(* IEC 61131-3 sources: RootPLC/conformance/cases/lexical, 40 files *)

(* ---- warn_soft_keyword_name.st ---- *)
(* spec: [lexical.keywords.soft]
   expect: warning RP0124
   run: PRG_Main cycles=2
   assert: n = 2
   assert: lit = TRUE *)
FUNCTION_BLOCK FB_Sequence
VAR_INPUT
    Step : INT;
    On : BOOL;
END_VAR
VAR_OUTPUT
    Task : DINT;
END_VAR
CASE Step OF
    1: Task := Task + 1;
END_CASE;
END_FUNCTION_BLOCK

PROGRAM PRG_Main
VAR
    seq : FB_Sequence;
    n : DINT;
    lit : BOOL;
    lamp AT %QX0.0 : BOOL;
END_VAR
seq(Step := 1, On := TRUE);
n := seq.Task;
lamp := seq.On;
lit := lamp;
END_PROGRAM

(* ---- err_bad_based_digit.st ---- *)
(* spec: [lexical.literal.integer]
   expect: error RP0008 *)
PROGRAM PRG_Main
VAR
    x : INT := 8#19;
END_VAR

END_PROGRAM

(* ---- err_bad_escape.st ---- *)
(* spec: [lexical.literal.escape]
   expect: error RP0010 *)
PROGRAM PRG_Main
VAR
    s : STRING := 'a$Qb';
END_VAR

END_PROGRAM

(* ---- err_char_two.st ---- *)
(* spec: [lexical.literal.char]
   expect: error RP0008 *)
PROGRAM PRG_Main
VAR
    c : CHAR := CHAR#'ab';
END_VAR

END_PROGRAM

(* ---- err_date_invalid.st ---- *)
(* spec: [lexical.literal.date]
   expect: error RP0012 *)
PROGRAM PRG_Main
VAR
    d : DATE := D#2026-02-30;
END_VAR

END_PROGRAM

(* ---- err_direct_variable.st ---- *)
(* spec: [lexical.direct-variable]
   expect: error RP0016 *)
PROGRAM PRG_Main
VAR
    x AT %IZ0 : BOOL;
END_VAR

END_PROGRAM

(* ---- err_duration_fraction_not_last.st ---- *)
(* spec: [lexical.literal.duration]
   expect: error RP0011 *)
PROGRAM PRG_Main
VAR
    t : TIME := T#1.5s20ms;
END_VAR

END_PROGRAM

(* ---- err_duration_order.st ---- *)
(* spec: [lexical.literal.duration]
   expect: error RP0011 *)
PROGRAM PRG_Main
VAR
    t : TIME := T#5s1m;
END_VAR

END_PROGRAM

(* ---- err_invalid_char.st ---- *)
(* spec: [lexical.source.charset] [lexical.punctuation]
   expect: error RP0005 *)
PROGRAM PRG_Main
VAR
    x : INT;
END_VAR
x := 1 @ 2;
END_PROGRAM

(* ---- err_keyword_identifier.st ---- *)
(* spec: [lexical.keyword]
   expect: error RP0004 *)
PROGRAM PRG_Main
VAR
    end_if : INT;
END_VAR

END_PROGRAM

(* ---- err_non_ascii_identifier.st ---- *)
(* spec: [lexical.source.charset]
   expect: error RP0005 *)
PROGRAM PRG_Main
VAR
    温度 : INT;
END_VAR

END_PROGRAM

(* ---- err_real_no_fraction.st ---- *)
(* spec: [lexical.literal.real]
   expect: error RP0008 *)
PROGRAM PRG_Main
VAR
    x : LREAL := 1.;
END_VAR

END_PROGRAM

(* ---- err_string_latin1.st ---- *)
(* spec: [lexical.literal.string.latin1]
   expect: error RP0009 *)
PROGRAM PRG_Main
VAR
    s : STRING := '温度';
END_VAR

END_PROGRAM

(* ---- err_tod_hour24.st ---- *)
(* spec: [lexical.literal.date]
   expect: error RP0012 *)
PROGRAM PRG_Main
VAR
    t : TOD := TOD#24:00:00;
END_VAR

END_PROGRAM

(* ---- err_typed_unknown.st ---- *)
(* spec: [lexical.literal.typed]
   expect: error RP0014 *)
PROGRAM PRG_Main
VAR
    x : INT := FOO#5;
END_VAR

END_PROGRAM

(* ---- err_underscore_double.st ---- *)
(* spec: [lexical.literal.underscore]
   expect: error RP0007 *)
PROGRAM PRG_Main
VAR
    x : INT := 1__0;
END_VAR

END_PROGRAM

(* ---- err_underscore_trailing.st ---- *)
(* spec: [lexical.literal.underscore]
   expect: error RP0007 *)
PROGRAM PRG_Main
VAR
    x : INT := 100_;
END_VAR

END_PROGRAM

(* ---- err_unterminated_comment.st ---- *)
(* spec: [lexical.comment.unterminated]
   expect: error RP0001 *)
PROGRAM PRG_Main (* never closed
END_PROGRAM

(* ---- err_unterminated_pragma.st ---- *)
(* spec: [lexical.pragma]
   expect: error RP0015 *)
PROGRAM PRG_Main
{attribute 'hide'
END_PROGRAM

(* ---- err_unterminated_string.st ---- *)
(* spec: [lexical.literal.string]
   expect: error RP0002 *)
PROGRAM PRG_Main
VAR
    s : STRING := 'abc
    n : INT;
END_VAR

END_PROGRAM

(* ---- ok_char_literals.st ---- *)
(* spec: [lexical.literal.char]
   expect: ok
   run: PRG_Main cycles=1
   assert: c = CHAR#'a' *)
PROGRAM PRG_Main
VAR
    c : CHAR := CHAR#'a';
    w : WCHAR := WCHAR#"b";
END_VAR

END_PROGRAM

(* ---- ok_comments.st ---- *)
(* spec: [lexical.comment.block] [lexical.comment.cblock] [lexical.comment.line] [lexical.whitespace] [lexical.source.encoding]
   expect: ok
   run: PRG_Main cycles=1
   assert: s = '/* not a comment */'
   assert: n = 1 *)
PROGRAM PRG_Main
VAR
    s : STRING := '/* not a comment */'; // line comment
    s2 : STRING := '(* not a comment *)';
	n : INT; /* C-style */
END_VAR
(* block
   comment *)
n := 1;
END_PROGRAM

(* ---- ok_date_literals.st ---- *)
(* spec: [lexical.literal.date]
   expect: ok *)
PROGRAM PRG_Main
VAR
    d : DATE := D#2026-11-03;
    t_day : TOD := TOD#14:30:00.5;
    stamp : DT := DT#2026-11-03-14:30:00;
    ld : LDATE := LDATE#2024-02-29;
END_VAR

END_PROGRAM

(* ---- ok_direct_variable.st ---- *)
(* spec: [lexical.direct-variable]
   expect: ok *)
PROGRAM PRG_Main
VAR
    start_btn AT %IX0.0 : BOOL;
    lamp AT %QX0.1 : BOOL;
    level AT %IW2 : WORD;
    spare AT %I* : BOOL;
END_VAR

END_PROGRAM

(* ---- ok_duration_literals.st ---- *)
(* spec: [lexical.literal.duration]
   expect: ok
   run: PRG_Main cycles=1
   assert: t1 = T#90m
   assert: t3 = T#1500ms *)
PROGRAM PRG_Main
VAR
    t1 : TIME := T#1h_30m;
    t2 : TIME := T#90m;
    t3 : TIME := T#1.5s;
    t4 : LTIME := LTIME#5us;
    t5 : TIME := t#-250ms;
END_VAR

END_PROGRAM

(* ---- ok_identifier_case.st ---- *)
(* spec: [lexical.identifier] [lexical.identifier.case]
   expect: ok
   run: PRG_Main cycles=1
   assert: motor_on = TRUE
   assert: _x1 = 3 *)
PROGRAM PRG_Main
VAR
    Motor_On : BOOL;
    _x1 : INT;
END_VAR
MOTOR_ON := TRUE;
_X1 := 3;
END_PROGRAM

(* ---- ok_integer_literals.st ---- *)
(* spec: [lexical.literal.integer] [lexical.literal.underscore] [lexical.literal.sign]
   expect: ok
   run: PRG_Main cycles=1
   assert: a = 1000000
   assert: b = 165
   assert: c = 15
   assert: d = 255
   assert: e = -128 *)
PROGRAM PRG_Main
VAR
    a : DINT := 1_000_000;
    b : INT := 2#1010_0101;
    c : INT := 8#17;
    d : DINT := 16#ff;
    e : SINT := -128;
END_VAR

END_PROGRAM

(* ---- ok_longest_match.st ---- *)
(* spec: [lexical.longest-match] [lexical.punctuation] [types.derived.array]
   expect: ok
   run: PRG_Main cycles=1
   assert: b = TRUE
   assert: a[10] = 1 *)
PROGRAM PRG_Main
VAR
    a : ARRAY[1..10] OF INT;
    x : INT := 1;
    y : INT := 2;
    b : BOOL;
END_VAR
b := x<=y;
a[10] := x**2;
END_PROGRAM

(* ---- ok_pragma_attribute.st ---- *)
(* spec: [lexical.pragma]
   expect: ok *)
PROGRAM PRG_Main
VAR
    {attribute 'hide'}
    x : INT;
END_VAR

END_PROGRAM

(* ---- ok_real_literals.st ---- *)
(* spec: [lexical.literal.real]
   expect: ok
   run: PRG_Main cycles=1
   assert: r = 1500.0
   assert: s = 0.25
   assert: t = 0.01 *)
PROGRAM PRG_Main
VAR
    r : LREAL := 1.5E3;
    s : REAL := 0.25;
    t : LREAL := 1.0e-2;
END_VAR

END_PROGRAM

(* ---- ok_strings.st ---- *)
(* spec: [lexical.literal.string] [lexical.literal.escape]
   expect: ok
   run: PRG_Main cycles=1
   assert: h = 'A' *)
PROGRAM PRG_Main
VAR
    s : STRING := 'it$'s $$5$N';
    w : WSTRING := "say $"hi$"";
    h : STRING := '$41';
END_VAR

END_PROGRAM

(* ---- ok_typed_literals.st ---- *)
(* spec: [lexical.literal.typed] [lexical.literal.bool]
   expect: ok
   run: PRG_Main cycles=1
   assert: a = 5
   assert: b = 255
   assert: c = TRUE
   assert: d = TRUE
   assert: e = 1.5 *)
PROGRAM PRG_Main
VAR
    a : INT := INT#5;
    b : BYTE := BYTE#16#FF;
    c : BOOL := BOOL#1;
    d : BOOL := TRUE;
    e : REAL := REAL#1.5;
END_VAR

END_PROGRAM

(* ---- ok_wstring_unicode.st ---- *)
(* spec: [lexical.literal.string] [lexical.source.charset]
   expect: ok *)
PROGRAM PRG_Main
VAR
    w : WSTRING := "温度";
END_VAR

END_PROGRAM

(* ---- warn_double_underscore.st ---- *)
(* spec: [lexical.identifier.underscore]
   expect: warning RP0006 *)
PROGRAM PRG_Main
VAR
    motor__on : BOOL;
END_VAR

END_PROGRAM

(* ---- warn_duration_inner_overflow.st ---- *)
(* spec: [lexical.literal.duration]
   expect: warning RP0128
   run: PRG_Main cycles=1
   assert: t = T#150m *)
PROGRAM PRG_Main
VAR
    t : TIME := T#1h90m;
END_VAR

END_PROGRAM

(* ---- warn_nested_comment.st ---- *)
(* spec: [lexical.comment.nesting]
   expect: warning RP0003 *)
PROGRAM PRG_Main
VAR
    x : INT;
END_VAR
(* outer (* inner *)
x := 1;
END_PROGRAM

(* ---- warn_null_ref_names.st ---- *)
(* spec: [lexical.keywords.soft]
   expect: warning RP0124
   run: PRG_Main cycles=1
   assert: k = 3
   assert: isNull = TRUE *)
TYPE E_DATA_STATE : (NULL, INIT, READY); END_TYPE
TYPE ST_X :
STRUCT
    Ref : INT;
END_STRUCT;
END_TYPE

PROGRAM PRG_Main
VAR
    s : E_DATA_STATE := E_DATA_STATE#NULL;
    x : ST_X;
    k : INT;
    isNull : BOOL;
END_VAR
x.Ref := 3;
k := x.Ref;
isNull := s = E_DATA_STATE#NULL;
END_PROGRAM

(* ---- warn_real_exponent_no_point.st ---- *)
(* spec: [lexical.literal.real]
   expect: warning RP0017
   run: PRG_Main cycles=1
   assert: x = 1000.0
   assert: y > 0.0 AND y < 0.000002 *)
PROGRAM PRG_Main
VAR
    x : LREAL := 1E3;
    y : LREAL := 1E-6;
END_VAR

END_PROGRAM

(* ---- warn_tod_without_seconds.st ---- *)
(* spec: [lexical.literal.date] [scope.vendor-forms]
   expect: warning RP0133
   run: PRG_Main cycles=1
   assert: same = TRUE
   assert: dsame = TRUE *)
PROGRAM PRG_Main
VAR
    a : TOD := TOD#12:00;
    d : DT := DT#2000-01-01-08:30;
    same, dsame : BOOL;
END_VAR
same := a = TOD#12:00:00;
dsame := d = DT#2000-01-01-08:30:00;
END_PROGRAM

(* ---- warn_unknown_pragma.st ---- *)
(* spec: [lexical.pragma]
   expect: warning RP0013 *)
PROGRAM PRG_Main
VAR
    {no_such_pragma 1}
    x : INT;
END_VAR

END_PROGRAM
